SUBAPPLICATION Uebung_264_AX (* RAMPO-Test: I1 = 8191, I2 = 0 auf Q1 RAMP 0ms, Q2 500ms, Q3 2s, Q4 Gamma 2s; je Ausgang CNF- und RAMPO-Zaehler *)
  (* Standard: 61499-2; Description: Copyright (c) 2026 Meisterschulen am Ostbahnhof This program and the accompanying materials are made available under the terms of the Eclipse Public License 2.0 which is available at https://www.eclipse.org/legal/epl-2.0/ SPDX-License-Identifier: EPL-2.0 *)
  (* Version 1.0, 2026-11-06, Franz Höpfinger, Meisterschulen am Ostbahnhof, initial API and implementation and/or initial documentation *)
  PACKAGE Uebungen;
  IMPORT logiBUS::io::DI::logiBUS_DI::Input_I1;
  IMPORT logiBUS::io::DI::logiBUS_DI::Input_I2;
  IMPORT logiBUS::io::DI::logiBUS_DI_Events::BUTTON_PRESS_DOWN;
  IMPORT logiBUS::io::DQ::logiBUS_DO::Output_Q1;
  IMPORT logiBUS::io::DQ::logiBUS_DO::Output_Q2;
  IMPORT logiBUS::io::DQ::logiBUS_DO::Output_Q3;
  IMPORT logiBUS::io::DQ::logiBUS_DO::Output_Q4;
  (* Documentation:
  RAMPO-Test
   I1 setzt 8191, I2 setzt 0. Q1 RAMP = T#0ms, Q2 T#500ms, Q3 T#2s, Q4 mit Gamma T#2s. Je Ausgang zählen CNF_Count_Qn und RAMPO_Count_Qn.
   Erwartung:
    - Ein neuer Wert: CNF +1, RAMPO +1 etwa nach der Rampenzeit (Q1 direkt nach dem CNF).
   - Zweimal schnell drücken: Q2 bis Q4 CNF +2, RAMPO +1 (die abgebrochene Rampe meldet kein RAMPO). Q1 springt jedes Mal: CNF +2, RAMPO +2.
   - Gleicher Taster zweimal (Ausgang steht schon auf dem Zielwert): keine Rampe, RAMPO kommt sofort, auch bei RAMP T#2s. Das ist richtig so.
   - Nach INIT kommt kein RAMPO.
    Kommt nie ein RAMPO oder stürzt die Firmware ab, passen Firmware und ELF nicht zusammen.
  *)
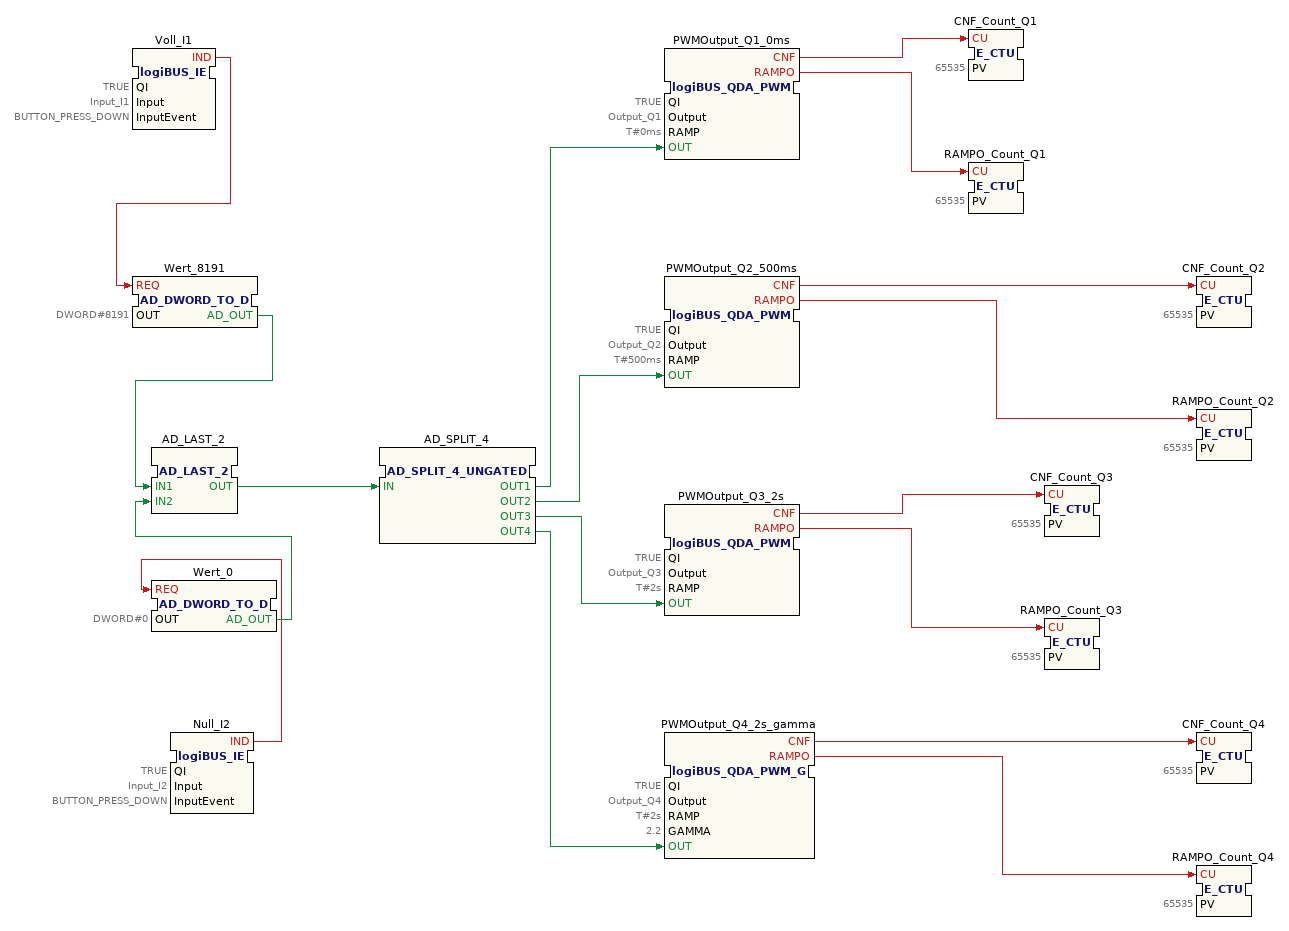
  FBS
    Voll_I1 : logiBUS::io::DI::logiBUS_IE(QI := TRUE, Input := Input_I1, InputEvent := BUTTON_PRESS_DOWN);
    Wert_8191 : adapter::conversion::unidirectional::AD_DWORD_TO_D(OUT := DWORD#8191);
    Null_I2 : logiBUS::io::DI::logiBUS_IE(QI := TRUE, Input := Input_I2, InputEvent := BUTTON_PRESS_DOWN);
    Wert_0 : adapter::conversion::unidirectional::AD_DWORD_TO_D(OUT := DWORD#0);
    AD_LAST_2 : adapter::events::unidirectional::AD_LAST_2;
    AD_SPLIT_4 : adapter::events::unidirectional::AD_SPLIT_4_UNGATED;
    PWMOutput_Q1_0ms : logiBUS::io::DQ::logiBUS_QDA_PWM(QI := TRUE, Output := Output_Q1, RAMP := T#0ms);
    CNF_Count_Q1 : iec61499::events::E_CTU(PV := 65535);
    RAMPO_Count_Q1 : iec61499::events::E_CTU(PV := 65535);
    PWMOutput_Q2_500ms : logiBUS::io::DQ::logiBUS_QDA_PWM(QI := TRUE, Output := Output_Q2, RAMP := T#500ms);
    CNF_Count_Q2 : iec61499::events::E_CTU(PV := 65535);
    RAMPO_Count_Q2 : iec61499::events::E_CTU(PV := 65535);
    PWMOutput_Q3_2s : logiBUS::io::DQ::logiBUS_QDA_PWM(QI := TRUE, Output := Output_Q3, RAMP := T#2s);
    CNF_Count_Q3 : iec61499::events::E_CTU(PV := 65535);
    RAMPO_Count_Q3 : iec61499::events::E_CTU(PV := 65535);
    PWMOutput_Q4_2s_gamma : logiBUS::io::DQ::logiBUS_QDA_PWM_G(QI := TRUE, Output := Output_Q4, RAMP := T#2s, GAMMA := 2.2);
    CNF_Count_Q4 : iec61499::events::E_CTU(PV := 65535);
    RAMPO_Count_Q4 : iec61499::events::E_CTU(PV := 65535);
  END_FBS
  EVENT_CONNECTIONS
    Voll_I1.IND TO Wert_8191.REQ;
    Null_I2.IND TO Wert_0.REQ;
    PWMOutput_Q1_0ms.CNF TO CNF_Count_Q1.CU;
    PWMOutput_Q1_0ms.RAMPO TO RAMPO_Count_Q1.CU;
    PWMOutput_Q2_500ms.CNF TO CNF_Count_Q2.CU;
    PWMOutput_Q2_500ms.RAMPO TO RAMPO_Count_Q2.CU;
    PWMOutput_Q3_2s.CNF TO CNF_Count_Q3.CU;
    PWMOutput_Q3_2s.RAMPO TO RAMPO_Count_Q3.CU;
    PWMOutput_Q4_2s_gamma.CNF TO CNF_Count_Q4.CU;
    PWMOutput_Q4_2s_gamma.RAMPO TO RAMPO_Count_Q4.CU;
  END_CONNECTIONS
  ADAPTER_CONNECTIONS
    Wert_8191.AD_OUT TO AD_LAST_2.IN1;
    Wert_0.AD_OUT TO AD_LAST_2.IN2;
    AD_LAST_2.OUT TO AD_SPLIT_4.IN;
    AD_SPLIT_4.OUT1 TO PWMOutput_Q1_0ms.OUT;
    AD_SPLIT_4.OUT2 TO PWMOutput_Q2_500ms.OUT;
    AD_SPLIT_4.OUT3 TO PWMOutput_Q3_2s.OUT;
    AD_SPLIT_4.OUT4 TO PWMOutput_Q4_2s_gamma.OUT;
  END_CONNECTIONS
END_SUBAPPLICATION
